Fanuc KAREL source: KT00864.KL

PROGRAM KT00864
%NOLOCKGROUP
VAR
  B1: BOOLEAN
  B2: BOOLEAN
  OUT: INTEGER
BEGIN
  B1 = TRUE
  B2 = FALSE
  B1 = TRUE
  B2 = FALSE
  OUT = ROUND(B1)
END KT00864
